Fanuc KAREL source: KT00732.KL

PROGRAM KT00732
%NOLOCKGROUP
VAR
  ARG: ARRAY[4] OF REAL
  OUT: BOOLEAN
BEGIN
  OUT = UNINIT(ARG)
END KT00732
